Fanuc KAREL source: compact_preamble.KL

PROGRAM KD00023
%NOLOCKGROUP
VAR
I:INTEGER;J:INTEGER;B:BOOLEAN;R:REAL;S : STRING[80];SAVED:INTEGER
BEGIN
I=SAVED
END KD00023
